// TIA Portal V20 export
TYPE "WT3_Feldbus_Header"
   STRUCT
      bKommAlarm { ExternalWritable := 'False'} : Bool;
      uiMbStartadresse { ExternalWritable := 'False'} : UInt;
      uiCount { S7_SetPoint := 'True'} : UInt;   // Anzahl WORD in Modbusdaten
      TON_Handshake : TON_TIME;
   END_STRUCT;
END_TYPE
